DATA_BLOCK "GDB_SequenceQuiesceTest"
{ S7_Optimized_Access := 'TRUE' }
VERSION : 0.1
NON_RETAIN
VAR
    Enabled : Bool;
    BeforeActive {ExternalWritable := 'False'} : Bool;
    AfterActive {ExternalWritable := 'False'} : Bool;
    HistorySurvived {ExternalWritable := 'False'} : Bool;
    CurrentCleared {ExternalWritable := 'False'} : Bool;
END_VAR
BEGIN
END_DATA_BLOCK
